// TIA Portal project "MiniProject_AziziFarid" (V16)

(* hardware
DEVICE "S71500/ET200MP station_1"  S7-1500 station
   slot 0: "Rail_0"  Rack  6ES7 590-1***0-0AA0
   slot 1: "AF_PLC_1 Distribution"  CPU 1512C-1 PN  6ES7 512-1CK00-0AB0  V2.6
      slot 3: "CPU display_1"  6ES7591-1AA00-0AA0
      slot 32768: "PROFINET interface_1"  X1
DEVICE "S71500/ET200MP station_2"  S7-1500 station
   slot 0: "Rail_0"  Rack  6ES7 590-1***0-0AA0
   slot 1: "AF_PLC_2 Joining"  CPU 1512C-1 PN  6ES7 512-1CK00-0AB0  V2.1
      slot 3: "CPU display_1"  6ES7591-1AA00-0AA0
      slot 32768: "PROFINET interface_1"  X1
DEVICE "S71500/ET200MP station_3"  S7-1500 station
   slot 0: "Rail_0"  Rack  6ES7 590-1***0-0AA0
   slot 1: "AF_PLC_3 Sorting"  CPU 1512C-1 PN  6ES7 512-1CK00-0AB0  V2.1
      slot 3: "CPU display_1"  6ES7591-1AA00-0AA0
      slot 32768: "PROFINET interface_1"  X1
DEVICE "GSD device_1"  GSD.Device.PN
   slot 0: "Rack"  Rack  V1.0
   slot 0: "CTEU-PN"  CTEU-PN  2201471
      slot 0: "CTEU-PN"  CTEU-PN
      slot 1: "PN-IO Interface"  PN-IO Interface
         slot 1: "Port 1"  Port 1
         slot 2: "Port 2"  Port 2
   slot 1: "Universal device 064DIO_1"  Universal device 064DIO
      slot 0: "Universal device 064DIO"  Universal device 064DIO
*)

// ===== PLC "AF_PLC_1 Distribution"  CPU 1512C-1 PN =====

VAR_GLOBAL   // PLC tag table "Default tag table"
   "SF1 START BTN" AT %I11.0 : Bool;
   "SF2 STOP BTN" AT %I11.1 : Bool;
   "SF4 KEY SWITCH" AT %I11.2 : Bool;
   "SF3 RESET BTN" AT %I11.3 : Bool;
   "G1BG1 SENSOR1" AT %I10.0 : Bool;
   "G1BG2 SENSOR2" AT %I10.1 : Bool;
   "G1BG3 SENSOR3" AT %I10.2 : Bool;
   "C2BG1 SLIDE RETRACT" AT %I10.4 : Bool;
   "C2BG2 SLIDE EXTEND" AT %I10.5 : Bool;
   "C2BG3 MAGAZINE EMPTY" AT %I10.6 : Bool;
   "PF1 START IND" AT %Q5.0 : Bool;
   "PF2 RESET IND" AT %Q5.1 : Bool;
   "PF3 IND Q1" AT %Q5.2 : Bool;
   "q4 XD4 STATION FREE" AT %Q5.4 : Bool;
   "q5 indLightGn" AT %Q5.5 : Bool;
   "q6 indLightYe" AT %Q5.6 : Bool;
   "q7 indLightRd" AT %Q5.7 : Bool;
   "G1BF1_A1 CONV FRWD" AT %Q4.0 : Bool;
   "G1BF1_A2 CONV BKWD" AT %Q4.1 : Bool;
   "G1MB1" AT %Q4.2 : Bool;
   "C2MB1" AT %Q4.4 : Bool;
   "System_Byte" AT %MB999 : Byte;
   "FirstScan" AT %M999.0 : Bool;
   "DiagStatusUpdate" AT %M999.1 : Bool;
   "AlwaysTRUE" AT %M999.2 : Bool;
   "AlwaysFALSE" AT %M999.3 : Bool;
   "Clock_Byte" AT %MB1000 : Byte;
   "Clock_10Hz" AT %M1000.0 : Bool;
   "Clock_5Hz" AT %M1000.1 : Bool;
   "Clock_2.5Hz" AT %M1000.2 : Bool;
   "Clock_2Hz" AT %M1000.3 : Bool;
   "Clock_1.25Hz" AT %M1000.4 : Bool;
   "Clock_1Hz" AT %M1000.5 : Bool;
   "Clock_0.625Hz" AT %M1000.6 : Bool;
   "Clock_0.5Hz" AT %M1000.7 : Bool;
   "xResetModules" AT %M200.0 : Bool;
   "xResetReadyModule1" AT %M200.1 : Bool;
   "xResetReadyModule2" AT %M200.2 : Bool;
   "xResetReadyModule3" AT %M200.3 : Bool;
   "xEnAutoMM" AT %M300.0 : Bool;
   "xDeactivateModules" AT %M200.6 : Bool;
   "xProcessBusyMM" AT %M200.7 : Bool;
   "xResetReadyMM" AT %M201.0 : Bool;
   "xNextStationFreeMM" AT %M201.1 : Bool;
   "xReadyModSM" AT %M201.2 : Bool;
   "xStartModuleSM" AT %M201.3 : Bool;
   "xMagEmptySM" AT %M201.4 : Bool;
   "xInitModules" AT %M201.5 : Bool;
   "PF4" AT %Q5.3 : Bool;
   "i7 XD7" AT %I11.7 : Bool;
   "i5 SF5" AT %I11.5 : Bool;
   "xResetReadyRFID_1" AT %M201.6 : Bool;
   "xMActivateModule1" AT %M201.7 : Bool;
   "xMEnAuto" AT %M400.7 : Bool;
   "xMStartProcess" AT %M300.2 : Bool;
   "xMProcessBusy" AT %M300.1 : Bool;
   "xMTP" AT %M203.0 : Bool;
   "xMTFR" AT %M203.1 : Bool;
   "xMG1BF1_A1" AT %M203.2 : Bool;
   "xM_MES_EnAuto" AT %M300.3 : Bool;
   "MWtest" AT %MW550 : Word;
   "bErrCodeMod1" AT %MB450 : Byte;
   "bErrCodeMod2" AT %MB451 : Byte;
   "bErrCodeMod3" AT %MB452 : Byte;
   "bErrCodeSeq" AT %MB453 : Byte;
   "bErrCodeOpMode" AT %MB454 : Byte;
   "Tag_1" AT %C2 : Counter;
   "i6 Jumper" AT %I11.6 : Bool;
   "Output" AT %M0.1 : Bool;
   "i4" AT %I11.4 : Bool;
   "Tag_2" AT %M0.0 : Bool;
   "Tag_3" AT %Q4.3 : Bool;
END_VAR

DATA_BLOCK "Dist_Block_DB"   // DB1
{ S7_Optimized_Access := 'TRUE' }
VERSION : 0.1
// stored: InstanceOfName Dist_Block
"Dist_Block"
BEGIN
END_DATA_BLOCK

// folder: System blocks/Program resources

DATA_BLOCK "IEC_Counter_0_DB"   // DB2
{ S7_Optimized_Access := 'TRUE' }
AUTHOR : Simatic
FAMILY : IEC
NAME : CNTR
VERSION : 1.0
// stored: InstanceOfName IEC_COUNTER
"IEC_COUNTER"
BEGIN
END_DATA_BLOCK

// folder: (top level)

FUNCTION_BLOCK "Dist_Block"   // FB2, GRAPH_PLUS
{ S7_Optimized_Access := 'TRUE' }
VERSION : 0.1
   VAR_INPUT
      OFF_SQ : Bool := false;   // Turn sequence off
      INIT_SQ : Bool := false;   // Set sequence to initial state
      ACK_EF : Bool := false;   // Acknowledge all errors and faults
      S_PREV : Bool := false;   // Output previous step in parameter S_NO
      S_NEXT : Bool := false;   // Indicate next step in parameter S_NO
      SW_AUTO : Bool := false;   // Automatic mode
      SW_TAP : Bool := false;   // Semiautomatic/switch with transition
      SW_TOP : Bool := false;   // Semiautomatic/ignore transition
      SW_MAN : Bool := false;   // Manual mode
      S_SEL : Int := 0;   // Select step to be output to S_NO
      S_ON : Bool := false;   // Activate step indicated in S_NO
      S_OFF : Bool := false;   // Deactivate step indicated S_NO
      T_PUSH : Bool := false;   // Enable transition to switch in semi automatic mode
   END_VAR
   VAR_OUTPUT
      S_NO : Int := 0;   // Step number
      S_MORE : Bool := false;   // More steps are available and can be shown in S_NO
      S_ACTIVE : Bool := false;   // Step indicated in S_NO is active
      ERR_FLT : Bool := false;   // Interlock or supervision group error
      AUTO_ON : Bool := false;   // Automatic mode is active
      TAP_ON : Bool := false;   // Semiautomatic mode/step with transition enabled
      TOP_ON : Bool := false;   // Semiautomatic mode/ignore transition enabled
      MAN_ON : Bool := false;   // Manual mode is active
   END_VAR
   VAR
      HMI_INFO : Array[0..8] of UInt;
      IF_PAR : G7_IfParPlus_V6;
      RT_DATA : G7_RTDataPlus_V6;   // Internal data area
      Trans1 : G7_TransitionPlus_V6;   // Transition structure
      Trans2 : G7_TransitionPlus_V6;   // Transition structure
      Trans3 : G7_TransitionPlus_V6;   // Transition structure
      Trans4 : G7_TransitionPlus_V6;   // Transition structure
      Trans5 : G7_TransitionPlus_V6;   // Transition structure
      Trans8 : G7_TransitionPlus_V6;   // Transition structure
      Trans9 : G7_TransitionPlus_V6;   // Transition structure
      Trans12 : G7_TransitionPlus_V6;   // Transition structure
      Trans13 : G7_TransitionPlus_V6;   // Transition structure
      Trans14 : G7_TransitionPlus_V6;   // Transition structure
      Step1 : G7_StepPlus_V6;   // Step structure
      Step2 : G7_StepPlus_V6;   // Step structure
      Step3 : G7_StepPlus_V6;   // Step structure
      Step4 : G7_StepPlus_V6;   // Step structure
      Step5 : G7_StepPlus_V6;   // Step structure
      Step8 : G7_StepPlus_V6;   // Step structure
      Step10 : G7_StepPlus_V6;   // Step structure
      Step11 : G7_StepPlus_V6;   // Step structure
      SINI : Array[0..1] of USInt;
      LSTT : Array[0..9] of USInt;
      ATAJ : Array[0..9] of USInt;
      ATAB : Array[0..9] of USInt;
      PSTT : Array[0..9] of USInt;
      NSTT : Array[0..9] of USInt;
      ASSJ : Array[0..7] of USInt;
      ASSB : Array[0..7] of USInt;
      PTTS : Array[0..7] of USInt;
      NTTS : Array[0..7] of USInt;
      SW_SQTS : Array[0..7] of USInt;
      SWITCH : Array[0..3] of USInt;
      TVX : Array[0..5] of USInt;
      TTX : Array[0..5] of USInt;
      TSX : Array[0..1] of USInt;
      S00X : Array[0..1] of USInt;
      SOFFX : Array[0..1] of USInt;
      SONX : Array[0..1] of USInt;
      SAX : Array[0..1] of USInt;
      SERRX : Array[0..8] of USInt;
      SMX : Array[0..8] of USInt;
      S0X : Array[0..8] of USInt;
      S1X : Array[0..8] of USInt;
      IL_ALARM_INST : Diag_Alarm;
      SUP_ALARM_INST : Diag_Alarm;
      STEP_TIME_ALARM_INST : Diag_Alarm;
      IEC_TIMER_INST : IEC_TIMER;
      TRANSACTION_FLAG : Bool := false;
   END_VAR
   // SINI[0] := 2;
   // LSTT[0] := 255;
   // LSTT[1] := 255;
   // LSTT[2] := 255;
   // ATAJ[1] := 1;
   // ATAJ[2] := 2;
   // ATAJ[3] := 3;
   // ATAB[1] := 1;
   // ATAB[2] := 2;
   // ATAB[3] := 7;
   // PSTT[1] := 1;
   // PSTT[2] := 2;
   // PSTT[3] := 3;
   // NSTT[0] := 1;
   // NSTT[1] := 2;
   // NSTT[2] := 3;
   // ASSJ[1] := 1;
   // ASSJ[2] := 2;
   // ASSJ[3] := 3;
   // ASSB[1] := 1;
   // ASSB[2] := 2;
   // ASSB[3] := 3;
   // PTTS[0] := 9;
   // PTTS[2] := 1;
   // PTTS[3] := 2;
   // NTTS[1] := 1;
   // NTTS[2] := 2;
   // NTTS[3] := 3;
   // TVX[0] := 16#1;
   // TTX[0] := 16#1;
   // TSX[0] := 16#1;
   // S00X[0] := 16#1;
   // SOFFX[0] := 16#1;
   // SONX[0] := 16#1;
   // SAX[0] := 16#1;
   // SERRX[0] := 16#1;
   // SMX[0] := 16#1;
   // S0X[0] := 16#1;
   // S1X[0] := 16#1;
   // ATAB[0] := 5;
   // LSTT[5] := 255;
   // ATAJ[4] := 4;
   // ATAJ[5] := 5;
   // ATAB[7] := 3;
   // NSTT[5] := 5;
   // ASSJ[4] := 4;
   // ASSB[4] := 4;
   // PTTS[4] := 3;
   // NTTS[4] := 4;
   // SW_SQTS[1] := 1;
   // SW_SQTS[2] := 1;
   // SW_SQTS[3] := 1;
   // SW_SQTS[4] := 2;
   // LSTT[3] := 255;
   // ATAJ[6] := 6;
   // ATAB[4] := 4;
   // PSTT[4] := 4;
   // NSTT[3] := 4;
   // ASSJ[5] := 5;
   // ASSB[5] := 5;
   // PTTS[5] := 5;
   // NTTS[6] := 8;
   // SW_SQTS[6] := 4;
   // LSTT[7] := 255;
   // ATAJ[7] := 7;
   // ATAB[6] := 6;
   // PSTT[7] := 3;
   // NSTT[7] := 6;
   // ASSJ[6] := 6;
   // ASSB[6] := 6;
   // PTTS[6] := 7;
   // NTTS[5] := 6;
   // LSTT[9] := 255;
   // ATAJ[8] := 8;
   // ATAJ[9] := 9;
   // ATAB[8] := 8;
   // ATAB[9] := 9;
   // PSTT[8] := 6;
   // PSTT[9] := 7;
   // ASSJ[7] := 7;
   // ASSB[7] := 7;
   // PTTS[7] := 255;
   // NTTS[7] := 9;
   // PSTT[6] := 5;
   // SW_SQTS[5] := 3;
BEGIN
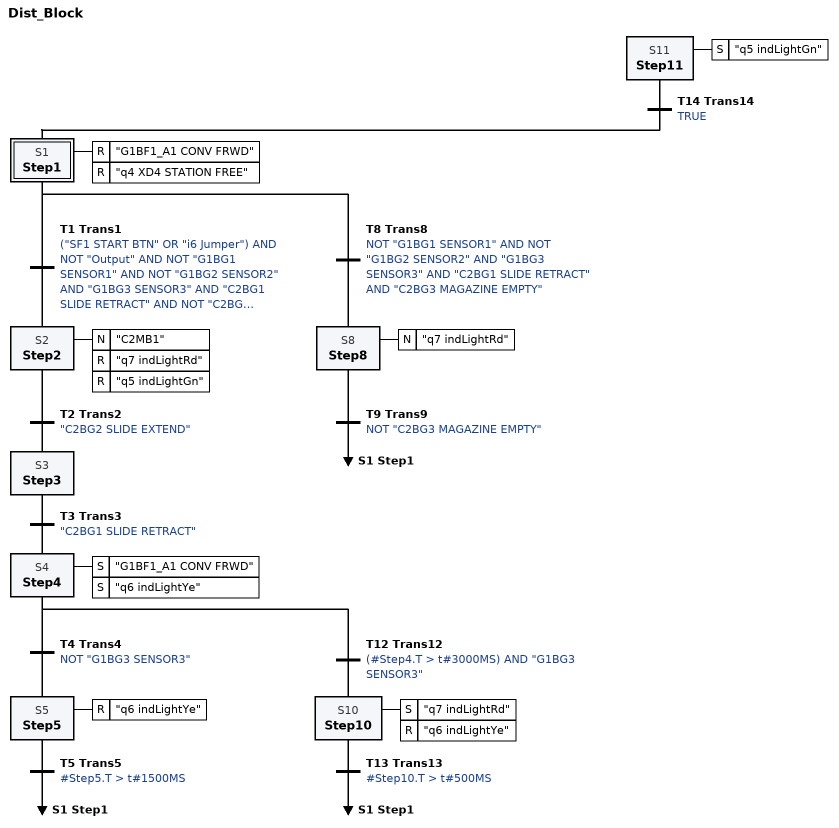
   // sequencer 1
   INITIAL_STEP Step1:   // S1, max time T#10S, warning time T#7S
              R    "G1BF1_A1 CONV FRWD"
              R    "q4 XD4 STATION FREE"
   END_STEP
   TRANSITION Trans1 FROM Step1 TO Step2   // T1
      := ("SF1 START BTN" OR "i6 Jumper") AND NOT "Output" AND NOT "G1BG1 SENSOR1" AND NOT "G1BG2 SENSOR2" AND "G1BG3 SENSOR3" AND "C2BG1 SLIDE RETRACT" AND NOT "C2BG3 MAGAZINE EMPTY";
   END_TRANSITION
   TRANSITION Trans8 FROM Step1 TO Step8   // T8
      := NOT "G1BG1 SENSOR1" AND NOT "G1BG2 SENSOR2" AND "G1BG3 SENSOR3" AND "C2BG1 SLIDE RETRACT" AND "C2BG3 MAGAZINE EMPTY";
   END_TRANSITION
   STEP Step2:   // S2, max time T#10S, warning time T#7S
              N    "C2MB1"
              R    "q7 indLightRd"
              R    "q5 indLightGn"
   END_STEP
   TRANSITION Trans2 FROM Step2 TO Step3   // T2
      := "C2BG2 SLIDE EXTEND";
   END_TRANSITION
   STEP Step3:   // S3, max time T#10S, warning time T#7S
   END_STEP
   TRANSITION Trans3 FROM Step3 TO Step4   // T3
      := "C2BG1 SLIDE RETRACT";
   END_TRANSITION
   STEP Step4:   // S4, max time T#10S, warning time T#7S
              S    "G1BF1_A1 CONV FRWD"
              S    "q6 indLightYe"
   END_STEP
   TRANSITION Trans4 FROM Step4 TO Step5   // T4
      := NOT "G1BG3 SENSOR3";
   END_TRANSITION
   TRANSITION Trans12 FROM Step4 TO Step10   // T12
      := (#Step4.T > t#3000MS) AND "G1BG3 SENSOR3";
   END_TRANSITION
   STEP Step8:   // S8, max time T#10S, warning time T#7S
              N    "q7 indLightRd"
   END_STEP
   TRANSITION Trans9 FROM Step8 TO Step1   // T9, jump
      := NOT "C2BG3 MAGAZINE EMPTY";
   END_TRANSITION
   STEP Step5:   // S5, max time T#10S, warning time T#7S
              R    "q6 indLightYe"
   END_STEP
   TRANSITION Trans5 FROM Step5 TO Step1   // T5, jump
      := #Step5.T > t#1500MS;
   END_TRANSITION
   STEP Step10:   // S10, max time T#10S, warning time T#7S
              S    "q7 indLightRd"
              R    "q6 indLightYe"
   END_STEP
   TRANSITION Trans13 FROM Step10 TO Step1   // T13, jump
      := #Step10.T > t#500MS;
   END_TRANSITION
   STEP Step11:   // S11, max time T#10S, warning time T#7S
              S    "q5 indLightGn"
   END_STEP
   TRANSITION Trans14 FROM Step11 TO Step1   // T14
      := TRUE;
   END_TRANSITION
END_FUNCTION_BLOCK

ORGANIZATION_BLOCK "Dist_Main"   // OB1, LAD, ProgramCycle
TITLE = "Main Program Sweep (Cycle)"
{ S7_Optimized_Access := 'TRUE' }
VERSION : 0.1
   VAR_INPUT
      Initial_Call : Bool;   // Initial call of this OB
      Remanence : Bool;   // =True, if remanent data are available
   END_VAR
BEGIN

REGION Network 1
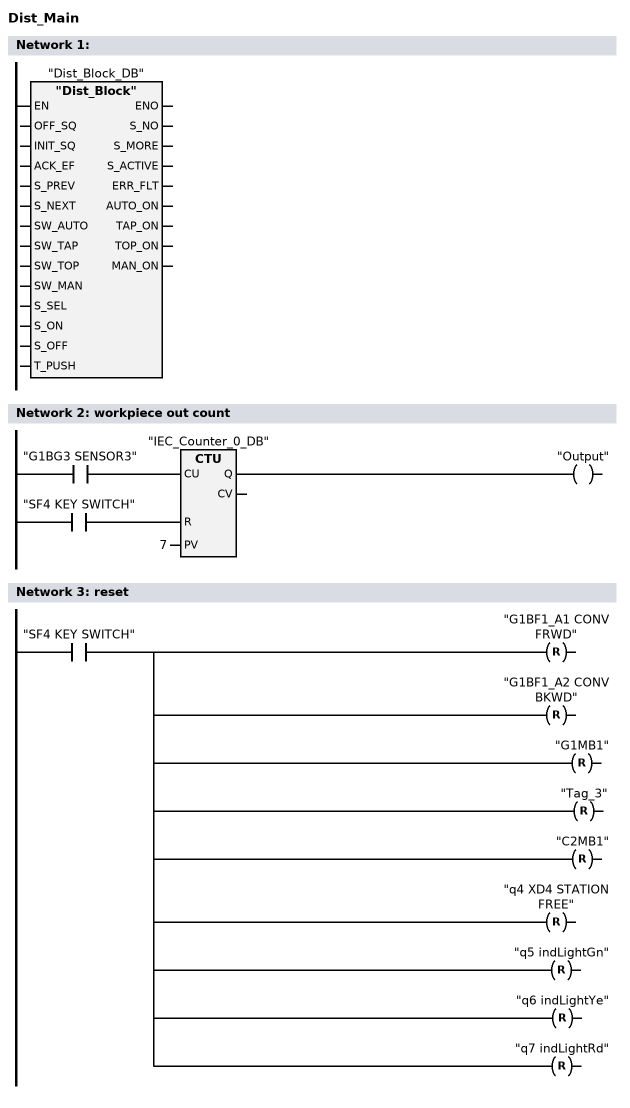
   RUNG wire#powerrail
      "Dist_Block_DB"(OFF_SQ :=, INIT_SQ :=, ACK_EF :=, S_PREV :=, S_NEXT :=, SW_AUTO :=, SW_TAP :=, SW_TOP :=, SW_MAN :=, S_SEL :=, S_ON :=, S_OFF :=, T_PUSH :=, S_NO =>, S_MORE =>, S_ACTIVE =>, ERR_FLT =>, AUTO_ON =>, TAP_ON =>, TOP_ON =>, MAN_ON =>)
   END_RUNG
   // the same network as SCL:
   "Dist_Block_DB"();   // "Dist_Block"
END_REGION

REGION Network 2: workpiece out count
   "IEC_Counter_0_DB".CTU(CU := "G1BG3 SENSOR3", R := "SF4 KEY SWITCH", PV := 7);
   "Output" := "IEC_Counter_0_DB".Q;
END_REGION

REGION Network 3: reset
   RUNG wire#powerrail
      Contact( "SF4 KEY SWITCH" )
      wire#w1
      R_Coil( "G1BF1_A1 CONV FRWD" )
   END_RUNG
   RUNG wire#w1
      R_Coil( "G1BF1_A2 CONV BKWD" )
   END_RUNG
   RUNG wire#w1
      R_Coil( "G1MB1" )
   END_RUNG
   RUNG wire#w1
      R_Coil( "Tag_3" )
   END_RUNG
   RUNG wire#w1
      R_Coil( "C2MB1" )
   END_RUNG
   RUNG wire#w1
      R_Coil( "q4 XD4 STATION FREE" )
   END_RUNG
   RUNG wire#w1
      R_Coil( "q5 indLightGn" )
   END_RUNG
   RUNG wire#w1
      R_Coil( "q6 indLightYe" )
   END_RUNG
   RUNG wire#w1
      R_Coil( "q7 indLightRd" )
   END_RUNG
   // the same network as SCL:
   IF "SF4 KEY SWITCH" THEN
       "G1BF1_A1 CONV FRWD" := FALSE;
       "G1BF1_A2 CONV BKWD" := FALSE;
       "G1MB1" := FALSE;
       "Tag_3" := FALSE;
       "C2MB1" := FALSE;
       "q4 XD4 STATION FREE" := FALSE;
       "q5 indLightGn" := FALSE;
       "q6 indLightYe" := FALSE;
       "q7 indLightRd" := FALSE;
   END_IF;
END_REGION
END_ORGANIZATION_BLOCK

// ===== PLC "AF_PLC_2 Joining"  CPU 1512C-1 PN =====

VAR_GLOBAL   // PLC tag table "Default tag table"
   "G1BG1 (diffuse 1 - depan)" AT %I10.0 : Bool;
   "G1BG2 (diffuse 2 - tengah)" AT %I10.1 : Bool;
   "G1MB1 (sep)" AT %Q4.2 : Bool;
   "G1MB2 (stopper)" AT %Q4.3 : Bool;
   "G1KF1-1 conv fwd" AT %Q4.0 : Bool;
   "G2BG3" AT %I10.6 : Bool;
   "G1KF1-2 conv bwd" AT %Q4.1 : Bool;
   "G1BG3 (through beam - hujung)" AT %I10.2 : Bool;
   "G1BG4 (distance)" AT %I10.3 : Bool;
   "G2KF1-1 conv fwd" AT %Q4.4 : Bool;
   "G2KF1-2 conv bwd" AT %Q4.5 : Bool;
   "G2BG1 (diffuse - capping)" AT %I10.4 : Bool;
   "SF1 (start btn)" AT %I11.0 : Bool;
   "SF2 (stop btn)" AT %I11.1 : Bool;
   "G3BG1 (sensor_arm_masuk)" AT %I126.0 : Bool;
   "G3BG2 (sensor_arm_keluar)" AT %I126.1 : Bool;
   "G3BG3 (sensor_arm_naik)" AT %I126.2 : Bool;
   "G3BP1 (sensor_sedut)" AT %I126.3 : Bool;
   "G3MB1 P1 (arm_keluar)" AT %Q128.1 : Bool;
   "G3MB2 P0 (arm_masuk)" AT %Q128.0 : Bool;
   "G3MB3 (arm_turunH_naikL)" AT %Q128.2 : Bool;
   "G3MB4 (sedut)" AT %Q128.3 : Bool;
   "SF3" AT %I11.2 : Bool;
   "SF4" AT %I11.3 : Bool;
   "i5" AT %I11.5 : Bool;
   "i6" AT %I11.6 : Bool;
   "i7" AT %I11.7 : Bool;
   "PF1" AT %I12.0 : Bool;
   "PF2" AT %I12.1 : Bool;
   "XPROCESSBUSY" AT %M0.0 : Bool;
   "i4 Jumper" AT %I11.4 : Bool;
   "output1" AT %M0.1 : Bool;
   "output2" AT %M0.2 : Bool;
   "q4" AT %Q5.4 : Bool;
   "q5" AT %Q5.5 : Bool;
   "q6" AT %Q5.6 : Bool;
   "q7" AT %Q5.7 : Bool;
END_VAR

DATA_BLOCK "Joining_Block_DB"   // DB1
{ S7_Optimized_Access := 'TRUE' }
VERSION : 0.1
// stored: InstanceOfName Joining_Block
"Joining_Block"
BEGIN
END_DATA_BLOCK

// folder: System blocks/Program resources

DATA_BLOCK "IEC_Counter_0_DB"   // DB2
{ S7_Optimized_Access := 'TRUE' }
AUTHOR : Simatic
FAMILY : IEC
NAME : CNTR
VERSION : 1.0
// stored: InstanceOfName IEC_COUNTER
"IEC_COUNTER"
BEGIN
END_DATA_BLOCK

DATA_BLOCK "IEC_Counter_0_DB_1"   // DB3
{ S7_Optimized_Access := 'TRUE' }
AUTHOR : Simatic
FAMILY : IEC
NAME : CNTR
VERSION : 1.0
// stored: InstanceOfName IEC_COUNTER
"IEC_COUNTER"
BEGIN
END_DATA_BLOCK

// folder: (top level)

FUNCTION_BLOCK "Joining_Block"   // FB1, GRAPH_PLUS
{ S7_Optimized_Access := 'TRUE' }
VERSION : 0.1
   VAR_INPUT
      OFF_SQ : Bool := false;   // Turn sequence off
      INIT_SQ : Bool := false;   // Set sequence to initial state
      ACK_EF : Bool := false;   // Acknowledge all errors and faults
      S_PREV : Bool := false;   // Output previous step in parameter S_NO
      S_NEXT : Bool := false;   // Indicate next step in parameter S_NO
      SW_AUTO : Bool := false;   // Automatic mode
      SW_TAP : Bool := false;   // Semiautomatic/switch with transition
      SW_TOP : Bool := false;   // Semiautomatic/ignore transition
      SW_MAN : Bool := false;   // Manual mode
      S_SEL : Int := 0;   // Select step to be output to S_NO
      S_ON : Bool := false;   // Activate step indicated in S_NO
      S_OFF : Bool := false;   // Deactivate step indicated S_NO
      T_PUSH : Bool := false;   // Enable transition to switch in semi automatic mode
   END_VAR
   VAR_OUTPUT
      S_NO : Int := 0;   // Step number
      S_MORE : Bool := false;   // More steps are available and can be shown in S_NO
      S_ACTIVE : Bool := false;   // Step indicated in S_NO is active
      ERR_FLT : Bool := false;   // Interlock or supervision group error
      AUTO_ON : Bool := false;   // Automatic mode is active
      TAP_ON : Bool := false;   // Semiautomatic mode/step with transition enabled
      TOP_ON : Bool := false;   // Semiautomatic mode/ignore transition enabled
      MAN_ON : Bool := false;   // Manual mode is active
   END_VAR
   VAR
      HMI_INFO : Array[0..8] of UInt;
      IF_PAR : G7_IfParPlus_V6;
      RT_DATA : G7_RTDataPlus_V6;   // Internal data area
      Trans1 : G7_TransitionPlus_V6;   // Transition structure
      Trans2 : G7_TransitionPlus_V6;   // Transition structure
      Trans3 : G7_TransitionPlus_V6;   // Transition structure
      Trans4 : G7_TransitionPlus_V6;   // Transition structure
      Trans5 : G7_TransitionPlus_V6;   // Transition structure
      Trans6 : G7_TransitionPlus_V6;   // Transition structure
      Trans7 : G7_TransitionPlus_V6;   // Transition structure
      Trans8 : G7_TransitionPlus_V6;   // Transition structure
      Trans9 : G7_TransitionPlus_V6;   // Transition structure
      Trans10 : G7_TransitionPlus_V6;   // Transition structure
      Trans11 : G7_TransitionPlus_V6;   // Transition structure
      Trans12 : G7_TransitionPlus_V6;   // Transition structure
      Trans13 : G7_TransitionPlus_V6;   // Transition structure
      Trans14 : G7_TransitionPlus_V6;   // Transition structure
      Trans15 : G7_TransitionPlus_V6;   // Transition structure
      Trans16 : G7_TransitionPlus_V6;   // Transition structure
      Trans17 : G7_TransitionPlus_V6;   // Transition structure
      Trans18 : G7_TransitionPlus_V6;   // Transition structure
      Trans19 : G7_TransitionPlus_V6;   // Transition structure
      Trans25 : G7_TransitionPlus_V6;   // Transition structure
      Trans26 : G7_TransitionPlus_V6;   // Transition structure
      Step1 : G7_StepPlus_V6;   // Step structure
      Step2 : G7_StepPlus_V6;   // Step structure
      Step3 : G7_StepPlus_V6;   // Step structure
      Step4 : G7_StepPlus_V6;   // Step structure
      Step5 : G7_StepPlus_V6;   // Step structure
      Step6 : G7_StepPlus_V6;   // Step structure
      Step8 : G7_StepPlus_V6;   // Step structure
      Step9 : G7_StepPlus_V6;   // Step structure
      Step10 : G7_StepPlus_V6;   // Step structure
      Step11 : G7_StepPlus_V6;   // Step structure
      Step12 : G7_StepPlus_V6;   // Step structure
      Step13 : G7_StepPlus_V6;   // Step structure
      Step14 : G7_StepPlus_V6;   // Step structure
      Step15 : G7_StepPlus_V6;   // Step structure
      Step16 : G7_StepPlus_V6;   // Step structure
      Step17 : G7_StepPlus_V6;   // Step structure
      Step18 : G7_StepPlus_V6;   // Step structure
      Step23 : G7_StepPlus_V6;   // Step structure
      Step24 : G7_StepPlus_V6;   // Step structure
      SINI : Array[0..1] of USInt;
      LSTT : Array[0..20] of USInt;
      ATAJ : Array[0..20] of USInt;
      ATAB : Array[0..20] of USInt;
      PSTT : Array[0..20] of USInt;
      NSTT : Array[0..20] of USInt;
      ASSJ : Array[0..18] of USInt;
      ASSB : Array[0..18] of USInt;
      PTTS : Array[0..18] of USInt;
      NTTS : Array[0..18] of USInt;
      SW_SQTS : Array[0..18] of USInt;
      SWITCH : Array[0..3] of USInt;
      TVX : Array[0..5] of USInt;
      TTX : Array[0..5] of USInt;
      TSX : Array[0..1] of USInt;
      S00X : Array[0..1] of USInt;
      SOFFX : Array[0..1] of USInt;
      SONX : Array[0..1] of USInt;
      SAX : Array[0..1] of USInt;
      SERRX : Array[0..19] of USInt;
      SMX : Array[0..19] of USInt;
      S0X : Array[0..19] of USInt;
      S1X : Array[0..19] of USInt;
      IL_ALARM_INST : Diag_Alarm;
      SUP_ALARM_INST : Diag_Alarm;
      STEP_TIME_ALARM_INST : Diag_Alarm;
      IEC_TIMER_INST : IEC_TIMER;
      TRANSACTION_FLAG : Bool := false;
   END_VAR
   // SINI[0] := 2;
   // LSTT[0] := 255;
   // LSTT[1] := 255;
   // LSTT[2] := 255;
   // LSTT[3] := 255;
   // LSTT[4] := 255;
   // LSTT[5] := 255;
   // LSTT[6] := 255;
   // LSTT[9] := 255;
   // ATAJ[1] := 1;
   // ATAJ[2] := 2;
   // ATAJ[3] := 3;
   // ATAJ[4] := 4;
   // ATAJ[5] := 5;
   // ATAJ[6] := 6;
   // ATAJ[7] := 7;
   // ATAJ[8] := 8;
   // ATAB[1] := 1;
   // ATAB[2] := 2;
   // ATAB[3] := 6;
   // ATAB[4] := 4;
   // ATAB[5] := 5;
   // ATAB[6] := 3;
   // ATAB[7] := 7;
   // ATAB[8] := 8;
   // PSTT[1] := 1;
   // PSTT[2] := 2;
   // PSTT[3] := 3;
   // PSTT[4] := 4;
   // PSTT[5] := 5;
   // PSTT[6] := 3;
   // PSTT[7] := 6;
   // PSTT[8] := 7;
   // NSTT[0] := 15;
   // NSTT[1] := 2;
   // NSTT[2] := 3;
   // NSTT[3] := 4;
   // NSTT[4] := 8;
   // NSTT[5] := 7;
   // NSTT[6] := 6;
   // NSTT[9] := 9;
   // ASSJ[1] := 1;
   // ASSJ[2] := 2;
   // ASSJ[3] := 3;
   // ASSJ[4] := 4;
   // ASSJ[5] := 5;
   // ASSJ[6] := 6;
   // ASSJ[7] := 7;
   // ASSB[1] := 1;
   // ASSB[2] := 2;
   // ASSB[3] := 3;
   // ASSB[4] := 4;
   // ASSB[5] := 5;
   // ASSB[6] := 6;
   // ASSB[7] := 7;
   // PTTS[0] := 255;
   // PTTS[2] := 1;
   // PTTS[3] := 2;
   // PTTS[4] := 3;
   // PTTS[5] := 14;
   // PTTS[6] := 6;
   // PTTS[7] := 5;
   // NTTS[1] := 1;
   // NTTS[2] := 2;
   // NTTS[3] := 3;
   // NTTS[4] := 4;
   // NTTS[5] := 5;
   // NTTS[6] := 7;
   // NTTS[7] := 8;
   // SW_SQTS[4] := 1;
   // SW_SQTS[5] := 2;
   // SW_SQTS[6] := 3;
   // SW_SQTS[7] := 2;
   // TVX[0] := 16#1;
   // TTX[0] := 16#1;
   // TSX[0] := 16#1;
   // S00X[0] := 16#1;
   // SOFFX[0] := 16#1;
   // SONX[0] := 16#1;
   // SAX[0] := 16#1;
   // SERRX[0] := 16#1;
   // SMX[0] := 16#1;
   // S0X[0] := 16#1;
   // S1X[0] := 16#1;
   // LSTT[10] := 255;
   // LSTT[11] := 255;
   // LSTT[12] := 255;
   // LSTT[13] := 255;
   // LSTT[14] := 255;
   // ATAJ[9] := 9;
   // ATAJ[10] := 10;
   // ATAJ[11] := 11;
   // ATAJ[12] := 12;
   // ATAJ[13] := 13;
   // ATAJ[14] := 14;
   // ATAB[9] := 9;
   // ATAB[10] := 17;
   // ATAB[11] := 11;
   // ATAB[12] := 12;
   // ATAB[13] := 13;
   // ATAB[14] := 14;
   // PSTT[9] := 8;
   // PSTT[10] := 9;
   // PSTT[11] := 10;
   // PSTT[12] := 11;
   // PSTT[13] := 12;
   // PSTT[14] := 13;
   // NSTT[10] := 10;
   // NSTT[11] := 11;
   // NSTT[12] := 12;
   // NSTT[13] := 13;
   // NSTT[14] := 5;
   // ASSJ[8] := 8;
   // ASSJ[9] := 9;
   // ASSJ[10] := 10;
   // ASSJ[11] := 11;
   // ASSJ[12] := 12;
   // ASSJ[13] := 13;
   // ASSB[8] := 8;
   // ASSB[9] := 9;
   // ASSB[10] := 10;
   // ASSB[11] := 11;
   // ASSB[12] := 12;
   // ASSB[13] := 13;
   // PTTS[8] := 4;
   // PTTS[9] := 9;
   // PTTS[10] := 10;
   // PTTS[11] := 11;
   // PTTS[12] := 12;
   // PTTS[13] := 13;
   // NTTS[8] := 9;
   // NTTS[9] := 10;
   // NTTS[10] := 11;
   // NTTS[11] := 12;
   // NTTS[12] := 13;
   // NTTS[13] := 14;
   // SW_SQTS[8] := 1;
   // SW_SQTS[9] := 1;
   // SW_SQTS[10] := 2;
   // SW_SQTS[11] := 2;
   // SW_SQTS[12] := 2;
   // SW_SQTS[13] := 2;
   // LSTT[7] := 255;
   // ATAJ[15] := 15;
   // ATAB[15] := 15;
   // PSTT[15] := 14;
   // NSTT[7] := 14;
   // ASSJ[14] := 14;
   // ASSB[14] := 14;
   // PTTS[14] := 7;
   // NTTS[14] := 15;
   // SW_SQTS[14] := 3;
   // LSTT[16] := 255;
   // ATAJ[16] := 16;
   // ATAB[16] := 16;
   // PSTT[16] := 15;
   // NSTT[16] := 1;
   // ASSJ[15] := 15;
   // ASSB[15] := 15;
   // PTTS[1] := 16;
   // NTTS[15] := 16;
   // LSTT[17] := 255;
   // LSTT[18] := 255;
   // ATAJ[17] := 17;
   // ATAJ[18] := 18;
   // ATAB[17] := 10;
   // ATAB[18] := 18;
   // PSTT[17] := 9;
   // PSTT[18] := 16;
   // NSTT[17] := 16;
   // NSTT[18] := 18;
   // ASSJ[16] := 16;
   // ASSB[16] := 16;
   // PTTS[16] := 17;
   // NTTS[16] := 18;
   // SW_SQTS[16] := 4;
   // LSTT[20] := 255;
   // ATAJ[19] := 19;
   // ATAJ[20] := 20;
   // ATAB[19] := 19;
   // ATAB[20] := 20;
   // PSTT[19] := 17;
   // PSTT[20] := 18;
   // NSTT[20] := 17;
   // ASSJ[17] := 17;
   // ASSJ[18] := 18;
   // ASSB[17] := 17;
   // ASSB[18] := 18;
   // PTTS[17] := 20;
   // PTTS[18] := 18;
   // NTTS[17] := 19;
   // NTTS[18] := 20;
   // SW_SQTS[17] := 4;
   // SW_SQTS[18] := 4;
BEGIN
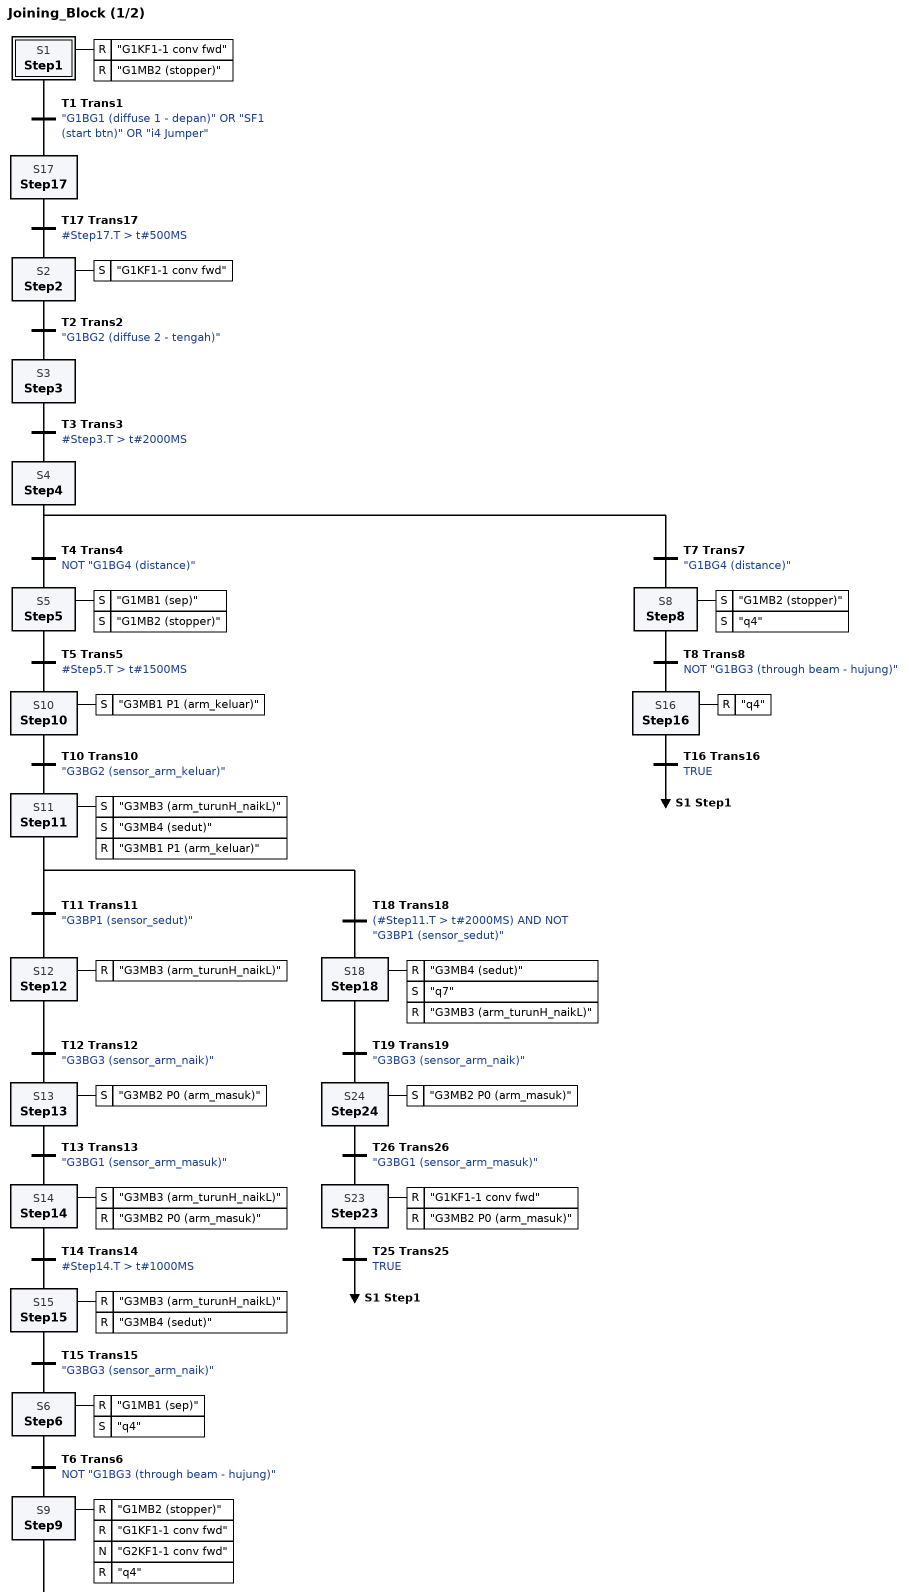
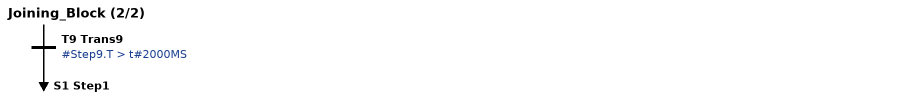
   // sequencer 1
   INITIAL_STEP Step1:   // S1, max time T#10S, warning time T#7S
              R    "G1KF1-1 conv fwd"
              R    "G1MB2 (stopper)"
   END_STEP
   TRANSITION Trans1 FROM Step1 TO Step17   // T1
      := "G1BG1 (diffuse 1 - depan)" OR "SF1 (start btn)" OR "i4 Jumper";
   END_TRANSITION
   STEP Step2:   // S2, max time T#10S, warning time T#7S
              S    "G1KF1-1 conv fwd"
   END_STEP
   TRANSITION Trans2 FROM Step2 TO Step3   // T2
      := "G1BG2 (diffuse 2 - tengah)";
   END_TRANSITION
   STEP Step3:   // S3, max time T#10S, warning time T#7S
   END_STEP
   TRANSITION Trans3 FROM Step3 TO Step4   // T3
      := #Step3.T > t#2000MS;
   END_TRANSITION
   STEP Step4:   // S4, max time T#10S, warning time T#7S
   END_STEP
   TRANSITION Trans4 FROM Step4 TO Step5   // T4
      := NOT "G1BG4 (distance)";
   END_TRANSITION
   TRANSITION Trans7 FROM Step4 TO Step8   // T7: Terbalik
      := "G1BG4 (distance)";
   END_TRANSITION
   STEP Step5:   // S5, max time T#10S, warning time T#7S
              S    "G1MB1 (sep)"
              S    "G1MB2 (stopper)"
   END_STEP
   TRANSITION Trans5 FROM Step5 TO Step10   // T5
      := #Step5.T > t#1500MS;
   END_TRANSITION
   STEP Step6:   // S6, max time T#10S, warning time T#7S
              R    "G1MB1 (sep)"
              S    "q4"
   END_STEP
   TRANSITION Trans6 FROM Step6 TO Step9   // T6
      := NOT "G1BG3 (through beam - hujung)";
   END_TRANSITION
   STEP Step8:   // S8, max time T#10S, warning time T#7S
              S    "G1MB2 (stopper)"
              S    "q4"
   END_STEP
   TRANSITION Trans8 FROM Step8 TO Step16   // T8
      := NOT "G1BG3 (through beam - hujung)";
   END_TRANSITION
   STEP Step9:   // S9, max time T#10S, warning time T#7S
              R    "G1MB2 (stopper)"
              R    "G1KF1-1 conv fwd"
              N    "G2KF1-1 conv fwd"
              R    "q4"
   END_STEP
   TRANSITION Trans9 FROM Step9 TO Step1   // T9, jump
      := #Step9.T > t#2000MS;
   END_TRANSITION
   STEP Step10:   // S10, max time T#10S, warning time T#7S
              S    "G3MB1 P1 (arm_keluar)"
   END_STEP
   TRANSITION Trans10 FROM Step10 TO Step11   // T10
      := "G3BG2 (sensor_arm_keluar)";
   END_TRANSITION
   STEP Step11:   // S11, max time T#10S, warning time T#7S
              S    "G3MB3 (arm_turunH_naikL)"
              S    "G3MB4 (sedut)"
              R    "G3MB1 P1 (arm_keluar)"
   END_STEP
   TRANSITION Trans11 FROM Step11 TO Step12   // T11
      := "G3BP1 (sensor_sedut)";
   END_TRANSITION
   TRANSITION Trans18 FROM Step11 TO Step18   // T18
      := (#Step11.T > t#2000MS) AND NOT "G3BP1 (sensor_sedut)";
   END_TRANSITION
   STEP Step12:   // S12, max time T#10S, warning time T#7S
              R    "G3MB3 (arm_turunH_naikL)"
   END_STEP
   TRANSITION Trans12 FROM Step12 TO Step13   // T12
      := "G3BG3 (sensor_arm_naik)";
   END_TRANSITION
   STEP Step13:   // S13, max time T#10S, warning time T#7S
      // undo Arm
              S    "G3MB2 P0 (arm_masuk)"
   END_STEP
   TRANSITION Trans13 FROM Step13 TO Step14   // T13
      := "G3BG1 (sensor_arm_masuk)";
   END_TRANSITION
   STEP Step14:   // S14, max time T#10S, warning time T#7S
      // turun Arm
              S    "G3MB3 (arm_turunH_naikL)"
              R    "G3MB2 P0 (arm_masuk)"
   END_STEP
   TRANSITION Trans14 FROM Step14 TO Step15   // T14
      := #Step14.T > t#1000MS;
   END_TRANSITION
   STEP Step15:   // S15, max time T#10S, warning time T#7S
      // pasang Cap
              R    "G3MB3 (arm_turunH_naikL)"
              R    "G3MB4 (sedut)"
   END_STEP
   TRANSITION Trans15 FROM Step15 TO Step6   // T15
      := "G3BG3 (sensor_arm_naik)";
   END_TRANSITION
   STEP Step16:   // S16, max time T#10S, warning time T#7S
              R    "q4"
   END_STEP
   TRANSITION Trans16 FROM Step16 TO Step1   // T16, jump
      := TRUE;
   END_TRANSITION
   STEP Step17:   // S17, max time T#10S, warning time T#7S
   END_STEP
   TRANSITION Trans17 FROM Step17 TO Step2   // T17
      := #Step17.T > t#500MS;
   END_TRANSITION
   STEP Step18:   // S18, max time T#10S, warning time T#7S
      // Lampu Merah
              R    "G3MB4 (sedut)"
              S    "q7"
              R    "G3MB3 (arm_turunH_naikL)"
   END_STEP
   TRANSITION Trans19 FROM Step18 TO Step24   // T19
      := "G3BG3 (sensor_arm_naik)";
   END_TRANSITION
   STEP Step24:   // S24, max time T#10S, warning time T#7S
              S    "G3MB2 P0 (arm_masuk)"
   END_STEP
   TRANSITION Trans26 FROM Step24 TO Step23   // T26
      := "G3BG1 (sensor_arm_masuk)";
   END_TRANSITION
   STEP Step23:   // S23, max time T#10S, warning time T#7S
              R    "G1KF1-1 conv fwd"
              R    "G3MB2 P0 (arm_masuk)"
   END_STEP
   TRANSITION Trans25 FROM Step23 TO Step1   // T25, jump
      := TRUE;
   END_TRANSITION
END_FUNCTION_BLOCK

ORGANIZATION_BLOCK "Joining_Main"   // OB1, LAD, ProgramCycle
TITLE = "Main Program Sweep (Cycle)"
{ S7_Optimized_Access := 'TRUE' }
VERSION : 0.1
   VAR_INPUT
      Initial_Call : Bool;   // Initial call of this OB
      Remanence : Bool;   // =True, if remanent data are available
   END_VAR
BEGIN

REGION Network 1
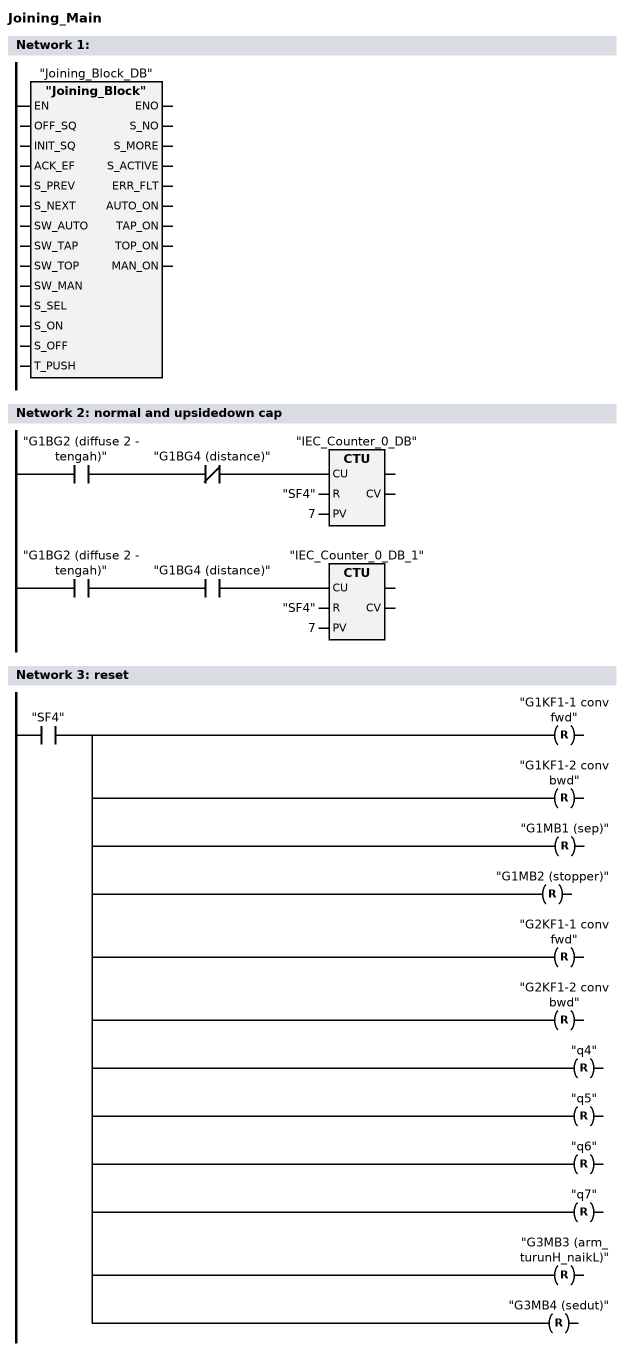
   RUNG wire#powerrail
      "Joining_Block_DB"(OFF_SQ :=, INIT_SQ :=, ACK_EF :=, S_PREV :=, S_NEXT :=, SW_AUTO :=, SW_TAP :=, SW_TOP :=, SW_MAN :=, S_SEL :=, S_ON :=, S_OFF :=, T_PUSH :=, S_NO =>, S_MORE =>, S_ACTIVE =>, ERR_FLT =>, AUTO_ON =>, TAP_ON =>, TOP_ON =>, MAN_ON =>)
   END_RUNG
   // the same network as SCL:
   "Joining_Block_DB"();   // "Joining_Block"
END_REGION

REGION Network 2: normal and upsidedown cap
   "IEC_Counter_0_DB".CTU(CU := "G1BG2 (diffuse 2 - tengah)" AND NOT "G1BG4 (distance)", R := "SF4", PV := 7);
   "IEC_Counter_0_DB_1".CTU(CU := "G1BG2 (diffuse 2 - tengah)" AND "G1BG4 (distance)", R := "SF4", PV := 7);
END_REGION

REGION Network 3: reset
   RUNG wire#powerrail
      Contact( "SF4" )
      wire#w1
      R_Coil( "G1KF1-1 conv fwd" )
   END_RUNG
   RUNG wire#w1
      R_Coil( "G1KF1-2 conv bwd" )
   END_RUNG
   RUNG wire#w1
      R_Coil( "G1MB1 (sep)" )
   END_RUNG
   RUNG wire#w1
      R_Coil( "G1MB2 (stopper)" )
   END_RUNG
   RUNG wire#w1
      R_Coil( "G2KF1-1 conv fwd" )
   END_RUNG
   RUNG wire#w1
      R_Coil( "G2KF1-2 conv bwd" )
   END_RUNG
   RUNG wire#w1
      R_Coil( "q4" )
   END_RUNG
   RUNG wire#w1
      R_Coil( "q5" )
   END_RUNG
   RUNG wire#w1
      R_Coil( "q6" )
   END_RUNG
   RUNG wire#w1
      R_Coil( "q7" )
   END_RUNG
   RUNG wire#w1
      R_Coil( "G3MB3 (arm_turunH_naikL)" )
   END_RUNG
   RUNG wire#w1
      R_Coil( "G3MB4 (sedut)" )
   END_RUNG
   // the same network as SCL:
   IF "SF4" THEN
       "G1KF1-1 conv fwd" := FALSE;
       "G1KF1-2 conv bwd" := FALSE;
       "G1MB1 (sep)" := FALSE;
       "G1MB2 (stopper)" := FALSE;
       "G2KF1-1 conv fwd" := FALSE;
       "G2KF1-2 conv bwd" := FALSE;
       "q4" := FALSE;
       "q5" := FALSE;
       "q6" := FALSE;
       "q7" := FALSE;
       "G3MB3 (arm_turunH_naikL)" := FALSE;
       "G3MB4 (sedut)" := FALSE;
   END_IF;
END_REGION
END_ORGANIZATION_BLOCK

// ===== PLC "AF_PLC_3 Sorting"  CPU 1512C-1 PN =====

VAR_GLOBAL   // PLC tag table "Default tag table"
   "SF1_START_BT" AT %I11.0 : Bool;
   "SF2_STOP_BT" AT %I11.1 : Bool;
   "SF4_KS MAN_AUTO" AT %I11.2 : Bool;
   "PF1_START INDI_LIGHT" AT %Q5.0 : Bool;
   "PF2_RESET INDI_LIGHT" AT %Q5.1 : Bool;
   "PF3(Q1)_INDI_LIGHT Q1" AT %Q5.2 : Bool;
   "PF4_INDI_LIGHT Q2" AT %Q5.3 : Bool;
   "B1BG1_FORK LIGHT BAR" AT %I10.4 : Bool;
   "B1BG2_RETRO LIGHT SENSOR" AT %I10.5 : Bool;
   "B1BG3_INDUC PROXI SENSOR" AT %I10.6 : Bool;
   "G1BG1_WP START" AT %I10.0 : Bool;
   "G1BG2_SEPARATOR 1 EXTRACT" AT %I10.1 : Bool;
   "G1BG4_SEPARATOR 2 EXTRACT" AT %I10.3 : Bool;
   "G1KF1_CONVEY MOTOR FOWD" AT %Q4.0 : Bool;
   "G1MB1_EXTEND SEPARATOR 1" AT %Q4.1 : Bool;
   "G1MB2_EXTEND SEPARATOR 2" AT %Q4.2 : Bool;
   "G1BG3_SENSOR SLIDE" AT %I10.2 : Bool;
   "G1MB3_RETRACT GATE" AT %Q4.3 : Bool;
   "q4 XD4_STATION FREE" AT %Q5.4 : Bool;
   "q5" AT %Q5.5 : Bool;
   "q6" AT %Q5.6 : Bool;
   "q7" AT %Q5.7 : Bool;
   "i4 Jumper" AT %I11.4 : Bool;
   "i5" AT %I11.5 : Bool;
   "i6 STATION_BUSY" AT %I11.6 : Bool;
   "i7" AT %I11.7 : Bool;
END_VAR

DATA_BLOCK "Sorting_Block_DB"   // DB1
{ S7_Optimized_Access := 'TRUE' }
VERSION : 0.1
// stored: InstanceOfName Sorting_Block
"Sorting_Block"
BEGIN
END_DATA_BLOCK

// folder: System blocks/Program resources

DATA_BLOCK "IEC_Counter_0_DB"   // DB2
{ S7_Optimized_Access := 'TRUE' }
AUTHOR : Simatic
FAMILY : IEC
NAME : CNTR
VERSION : 1.0
// stored: InstanceOfName IEC_COUNTER
"IEC_COUNTER"
BEGIN
END_DATA_BLOCK

DATA_BLOCK "IEC_Counter_0_DB_1"   // DB3
{ S7_Optimized_Access := 'TRUE' }
AUTHOR : Simatic
FAMILY : IEC
NAME : CNTR
VERSION : 1.0
// stored: InstanceOfName IEC_COUNTER
"IEC_COUNTER"
BEGIN
END_DATA_BLOCK

DATA_BLOCK "IEC_Counter_0_DB_2"   // DB4
{ S7_Optimized_Access := 'TRUE' }
AUTHOR : Simatic
FAMILY : IEC
NAME : CNTR
VERSION : 1.0
// stored: InstanceOfName IEC_COUNTER
"IEC_COUNTER"
BEGIN
END_DATA_BLOCK

// folder: (top level)

FUNCTION_BLOCK "Sorting_Block"   // FB3, GRAPH_PLUS
{ S7_Optimized_Access := 'TRUE' }
VERSION : 0.1
   VAR_INPUT
      OFF_SQ : Bool := false;   // Turn sequence off
      INIT_SQ : Bool := false;   // Set sequence to initial state
      ACK_EF : Bool := false;   // Acknowledge all errors and faults
      S_PREV : Bool := false;   // Output previous step in parameter S_NO
      S_NEXT : Bool := false;   // Indicate next step in parameter S_NO
      SW_AUTO : Bool := false;   // Automatic mode
      SW_TAP : Bool := false;   // Semiautomatic/switch with transition
      SW_TOP : Bool := false;   // Semiautomatic/ignore transition
      SW_MAN : Bool := false;   // Manual mode
      S_SEL : Int := 0;   // Select step to be output to S_NO
      S_ON : Bool := false;   // Activate step indicated in S_NO
      S_OFF : Bool := false;   // Deactivate step indicated S_NO
      T_PUSH : Bool := false;   // Enable transition to switch in semi automatic mode
   END_VAR
   VAR_OUTPUT
      S_NO : Int := 0;   // Step number
      S_MORE : Bool := false;   // More steps are available and can be shown in S_NO
      S_ACTIVE : Bool := false;   // Step indicated in S_NO is active
      ERR_FLT : Bool := false;   // Interlock or supervision group error
      AUTO_ON : Bool := false;   // Automatic mode is active
      TAP_ON : Bool := false;   // Semiautomatic mode/step with transition enabled
      TOP_ON : Bool := false;   // Semiautomatic mode/ignore transition enabled
      MAN_ON : Bool := false;   // Manual mode is active
   END_VAR
   VAR
      HMI_INFO : Array[0..8] of UInt;
      IF_PAR : G7_IfParPlus_V6;
      RT_DATA : G7_RTDataPlus_V6;   // Internal data area
      Trans1 : G7_TransitionPlus_V6;   // Transition structure
      Trans2 : G7_TransitionPlus_V6;   // Transition structure
      Trans3 : G7_TransitionPlus_V6;   // Transition structure
      Trans4 : G7_TransitionPlus_V6;   // Transition structure
      Trans5 : G7_TransitionPlus_V6;   // Transition structure
      Trans6 : G7_TransitionPlus_V6;   // Transition structure
      Trans7 : G7_TransitionPlus_V6;   // Transition structure
      Trans8 : G7_TransitionPlus_V6;   // Transition structure
      Trans9 : G7_TransitionPlus_V6;   // Transition structure
      Trans10 : G7_TransitionPlus_V6;   // Transition structure
      Trans11 : G7_TransitionPlus_V6;   // Transition structure
      Trans13 : G7_TransitionPlus_V6;   // Transition structure
      Trans14 : G7_TransitionPlus_V6;   // Transition structure
      Trans16 : G7_TransitionPlus_V6;   // Transition structure
      Trans17 : G7_TransitionPlus_V6;   // Transition structure
      Trans19 : G7_TransitionPlus_V6;   // Transition structure
      Trans20 : G7_TransitionPlus_V6;   // Transition structure
      Trans21 : G7_TransitionPlus_V6;   // Transition structure
      Step1 : G7_StepPlus_V6;   // Step structure
      Step2 : G7_StepPlus_V6;   // Step structure
      Step3 : G7_StepPlus_V6;   // Step structure
      Step4 : G7_StepPlus_V6;   // Step structure
      Step5 : G7_StepPlus_V6;   // Step structure
      Step6 : G7_StepPlus_V6;   // Step structure
      Step8 : G7_StepPlus_V6;   // Step structure
      Step9 : G7_StepPlus_V6;   // Step structure
      Step10 : G7_StepPlus_V6;   // Step structure
      Step12 : G7_StepPlus_V6;   // Step structure
      Step13 : G7_StepPlus_V6;   // Step structure
      Step14 : G7_StepPlus_V6;   // Step structure
      Step15 : G7_StepPlus_V6;   // Step structure
      Step16 : G7_StepPlus_V6;   // Step structure
      SINI : Array[0..1] of USInt;
      LSTT : Array[0..17] of USInt;
      ATAJ : Array[0..17] of USInt;
      ATAB : Array[0..17] of USInt;
      PSTT : Array[0..17] of USInt;
      NSTT : Array[0..17] of USInt;
      ASSJ : Array[0..13] of USInt;
      ASSB : Array[0..13] of USInt;
      PTTS : Array[0..13] of USInt;
      NTTS : Array[0..13] of USInt;
      SW_SQTS : Array[0..13] of USInt;
      SWITCH : Array[0..10] of USInt;
      TVX : Array[0..8] of USInt;
      TTX : Array[0..8] of USInt;
      TSX : Array[0..1] of USInt;
      S00X : Array[0..1] of USInt;
      SOFFX : Array[0..1] of USInt;
      SONX : Array[0..1] of USInt;
      SAX : Array[0..1] of USInt;
      SERRX : Array[0..14] of USInt;
      SMX : Array[0..14] of USInt;
      S0X : Array[0..14] of USInt;
      S1X : Array[0..14] of USInt;
      IL_ALARM_INST : Diag_Alarm;
      SUP_ALARM_INST : Diag_Alarm;
      STEP_TIME_ALARM_INST : Diag_Alarm;
      IEC_TIMER_INST : IEC_TIMER;
      TRANSACTION_FLAG : Bool := false;
   END_VAR
   // LSTT[13] := 255;
   // SINI[0] := 2;
   // LSTT[0] := 255;
   // LSTT[1] := 255;
   // LSTT[2] := 255;
   // LSTT[3] := 255;
   // LSTT[4] := 255;
   // LSTT[5] := 255;
   // LSTT[6] := 255;
   // LSTT[7] := 255;
   // LSTT[8] := 255;
   // LSTT[9] := 255;
   // LSTT[10] := 255;
   // ATAJ[1] := 1;
   // ATAJ[2] := 2;
   // ATAJ[3] := 3;
   // ATAJ[4] := 4;
   // ATAJ[5] := 6;
   // ATAJ[6] := 10;
   // ATAJ[7] := 7;
   // ATAJ[8] := 8;
   // ATAJ[9] := 9;
   // ATAJ[10] := 5;
   // ATAJ[11] := 11;
   // ATAJ[12] := 12;
   // ATAB[0] := 1;
   // ATAB[1] := 2;
   // ATAB[3] := 12;
   // ATAB[4] := 15;
   // ATAB[5] := 5;
   // ATAB[6] := 6;
   // ATAB[7] := 7;
   // ATAB[8] := 8;
   // ATAB[9] := 9;
   // ATAB[10] := 10;
   // ATAB[11] := 11;
   // ATAB[12] := 3;
   // PSTT[0] := 8;
   // PSTT[1] := 8;
   // PSTT[2] := 8;
   // PSTT[3] := 1;
   // PSTT[4] := 2;
   // PSTT[5] := 3;
   // PSTT[6] := 4;
   // PSTT[8] := 6;
   // PSTT[9] := 7;
   // PSTT[10] := 5;
   // PSTT[11] := 10;
   // PSTT[12] := 1;
   // NSTT[13] := 11;
   // NSTT[0] := 1;
   // NSTT[1] := 2;
   // NSTT[2] := 3;
   // NSTT[3] := 4;
   // NSTT[4] := 5;
   // NSTT[5] := 10;
   // NSTT[6] := 10;
   // NSTT[7] := 6;
   // NSTT[8] := 7;
   // NSTT[9] := 8;
   // NSTT[10] := 10;
   // ASSJ[1] := 1;
   // ASSJ[2] := 2;
   // ASSJ[3] := 3;
   // ASSJ[4] := 4;
   // ASSJ[5] := 5;
   // ASSJ[6] := 6;
   // ASSJ[7] := 7;
   // ASSJ[8] := 8;
   // ASSJ[9] := 9;
   // ASSJ[10] := 10;
   // ASSB[1] := 1;
   // ASSB[2] := 2;
   // ASSB[3] := 3;
   // ASSB[4] := 4;
   // ASSB[5] := 5;
   // ASSB[6] := 6;
   // ASSB[7] := 7;
   // ASSB[8] := 8;
   // ASSB[9] := 9;
   // ASSB[10] := 10;
   // PTTS[0] := 255;
   // PTTS[2] := 1;
   // PTTS[3] := 2;
   // PTTS[4] := 3;
   // PTTS[5] := 4;
   // PTTS[6] := 7;
   // PTTS[7] := 8;
   // PTTS[8] := 9;
   // PTTS[9] := 12;
   // PTTS[10] := 6;
   // NTTS[0] := 7;
   // NTTS[1] := 3;
   // NTTS[2] := 4;
   // NTTS[3] := 5;
   // NTTS[4] := 6;
   // NTTS[5] := 10;
   // NTTS[6] := 8;
   // NTTS[7] := 9;
   // NTTS[9] := 13;
   // NTTS[10] := 11;
   // SW_SQTS[1] := 1;
   // SW_SQTS[2] := 2;
   // SW_SQTS[3] := 3;
   // SW_SQTS[4] := 4;
   // SW_SQTS[5] := 5;
   // SW_SQTS[9] := 6;
   // SW_SQTS[10] := 7;
   // TVX[0] := 16#1;
   // TTX[0] := 16#1;
   // TSX[0] := 16#1;
   // S00X[0] := 16#1;
   // SOFFX[0] := 16#1;
   // SONX[0] := 16#1;
   // SAX[0] := 16#1;
   // SERRX[0] := 16#1;
   // SMX[0] := 16#1;
   // S0X[0] := 16#1;
   // S1X[0] := 16#1;
   // LSTT[12] := 255;
   // LSTT[14] := 4;
   // LSTT[15] := 255;
   // ATAJ[13] := 13;
   // ATAJ[14] := 14;
   // ATAJ[15] := 15;
   // ATAB[13] := 13;
   // ATAB[14] := 14;
   // ATAB[15] := 4;
   // PSTT[13] := 9;
   // PSTT[14] := 11;
   // PSTT[15] := 2;
   // NSTT[12] := 9;
   // NSTT[14] := 4;
   // NSTT[15] := 12;
   // ASSJ[11] := 11;
   // ASSJ[12] := 12;
   // ASSB[11] := 11;
   // ASSB[12] := 12;
   // PTTS[11] := 13;
   // PTTS[12] := 15;
   // NTTS[11] := 14;
   // NTTS[12] := 16;
   // SW_SQTS[11] := 6;
   // SW_SQTS[12] := 8;
   // LSTT[16] := 255;
   // LSTT[17] := 4;
   // ATAJ[16] := 16;
   // ATAJ[17] := 17;
   // ATAB[16] := 16;
   // ATAB[17] := 17;
   // PSTT[16] := 12;
   // PSTT[17] := 13;
   // NSTT[16] := 13;
   // NSTT[17] := 4;
   // ASSJ[13] := 13;
   // ASSB[13] := 13;
   // PTTS[13] := 16;
   // NTTS[13] := 17;
   // SW_SQTS[13] := 8;
BEGIN
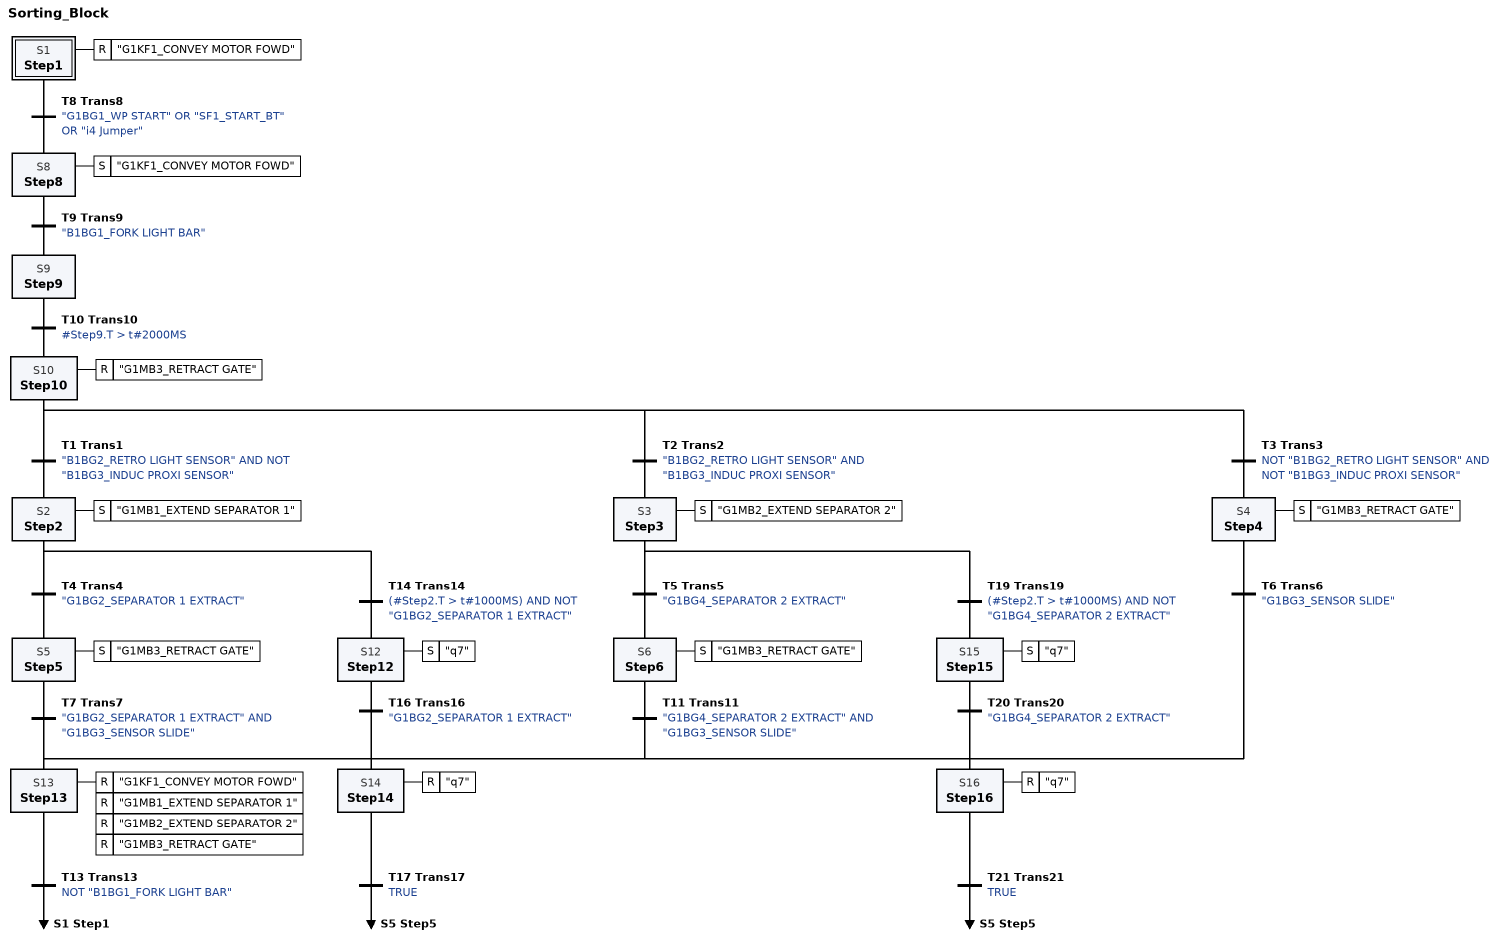
   // sequencer 1
   INITIAL_STEP Step1:   // S1, max time T#10S, warning time T#7S
              R    "G1KF1_CONVEY MOTOR FOWD"
   END_STEP
   TRANSITION Trans8 FROM Step1 TO Step8   // T8
      := "G1BG1_WP START" OR "SF1_START_BT" OR "i4 Jumper";
   END_TRANSITION
   STEP Step2:   // S2, max time T#10S, warning time T#7S
              S    "G1MB1_EXTEND SEPARATOR 1"
   END_STEP
   TRANSITION Trans4 FROM Step2 TO Step5   // T4
      := "G1BG2_SEPARATOR 1 EXTRACT";
   END_TRANSITION
   TRANSITION Trans14 FROM Step2 TO Step12   // T14
      := (#Step2.T > t#1000MS) AND NOT "G1BG2_SEPARATOR 1 EXTRACT";
   END_TRANSITION
   STEP Step3:   // S3, max time T#10S, warning time T#7S
              S    "G1MB2_EXTEND SEPARATOR 2"
   END_STEP
   TRANSITION Trans5 FROM Step3 TO Step6   // T5
      := "G1BG4_SEPARATOR 2 EXTRACT";
   END_TRANSITION
   TRANSITION Trans19 FROM Step3 TO Step15   // T19
      := (#Step2.T > t#1000MS) AND NOT "G1BG4_SEPARATOR 2 EXTRACT";
   END_TRANSITION
   STEP Step4:   // S4, max time T#10S, warning time T#7S
              S    "G1MB3_RETRACT GATE"
   END_STEP
   TRANSITION Trans6 FROM Step4 TO Step13   // T6
      := "G1BG3_SENSOR SLIDE";
   END_TRANSITION
   STEP Step5:   // S5, max time T#10S, warning time T#7S
              S    "G1MB3_RETRACT GATE"
   END_STEP
   TRANSITION Trans7 FROM Step5 TO Step13   // T7
      := "G1BG2_SEPARATOR 1 EXTRACT" AND "G1BG3_SENSOR SLIDE";
   END_TRANSITION
   STEP Step6:   // S6, max time T#10S, warning time T#7S
              S    "G1MB3_RETRACT GATE"
   END_STEP
   TRANSITION Trans11 FROM Step6 TO Step13   // T11
      := "G1BG4_SEPARATOR 2 EXTRACT" AND "G1BG3_SENSOR SLIDE";
   END_TRANSITION
   STEP Step8:   // S8, max time T#10S, warning time T#7S
              S    "G1KF1_CONVEY MOTOR FOWD"
   END_STEP
   TRANSITION Trans9 FROM Step8 TO Step9   // T9
      := "B1BG1_FORK LIGHT BAR";
   END_TRANSITION
   STEP Step10:   // S10, max time T#10S, warning time T#7S
              R    "G1MB3_RETRACT GATE"
   END_STEP
   TRANSITION Trans1 FROM Step10 TO Step2   // T1
      := "B1BG2_RETRO LIGHT SENSOR" AND NOT "B1BG3_INDUC PROXI SENSOR";
   END_TRANSITION
   TRANSITION Trans2 FROM Step10 TO Step3   // T2
      := "B1BG2_RETRO LIGHT SENSOR" AND "B1BG3_INDUC PROXI SENSOR";
   END_TRANSITION
   TRANSITION Trans3 FROM Step10 TO Step4   // T3
      := NOT "B1BG2_RETRO LIGHT SENSOR" AND NOT "B1BG3_INDUC PROXI SENSOR";
   END_TRANSITION
   STEP Step9:   // S9, max time T#10S, warning time T#7S
   END_STEP
   TRANSITION Trans10 FROM Step9 TO Step10   // T10
      := #Step9.T > t#2000MS;
   END_TRANSITION
   STEP Step12:   // S12, max time T#10S, warning time T#7S
              S    "q7"
   END_STEP
   TRANSITION Trans16 FROM Step12 TO Step14   // T16
      := "G1BG2_SEPARATOR 1 EXTRACT";
   END_TRANSITION
   STEP Step14:   // S14, max time T#10S, warning time T#7S
              R    "q7"
   END_STEP
   TRANSITION Trans17 FROM Step14 TO Step5   // T17, jump
      := TRUE;
   END_TRANSITION
   STEP Step15:   // S15, max time T#10S, warning time T#7S
              S    "q7"
   END_STEP
   TRANSITION Trans20 FROM Step15 TO Step16   // T20
      := "G1BG4_SEPARATOR 2 EXTRACT";
   END_TRANSITION
   STEP Step16:   // S16, max time T#10S, warning time T#7S
              R    "q7"
   END_STEP
   TRANSITION Trans21 FROM Step16 TO Step5   // T21, jump
      := TRUE;
   END_TRANSITION
   STEP Step13:   // S13, max time T#10S, warning time T#7S
              R    "G1KF1_CONVEY MOTOR FOWD"
              R    "G1MB1_EXTEND SEPARATOR 1"
              R    "G1MB2_EXTEND SEPARATOR 2"
              R    "G1MB3_RETRACT GATE"
   END_STEP
   TRANSITION Trans13 FROM Step13 TO Step1   // T13, jump
      := NOT "B1BG1_FORK LIGHT BAR";
   END_TRANSITION
END_FUNCTION_BLOCK

ORGANIZATION_BLOCK "Sorting_Main"   // OB1, LAD, ProgramCycle
TITLE = "Main Program Sweep (Cycle)"
{ S7_Optimized_Access := 'TRUE' }
VERSION : 0.1
   VAR_INPUT
      Initial_Call : Bool;   // Initial call of this OB
      Remanence : Bool;   // =True, if remanent data are available
   END_VAR
BEGIN

REGION Network 1
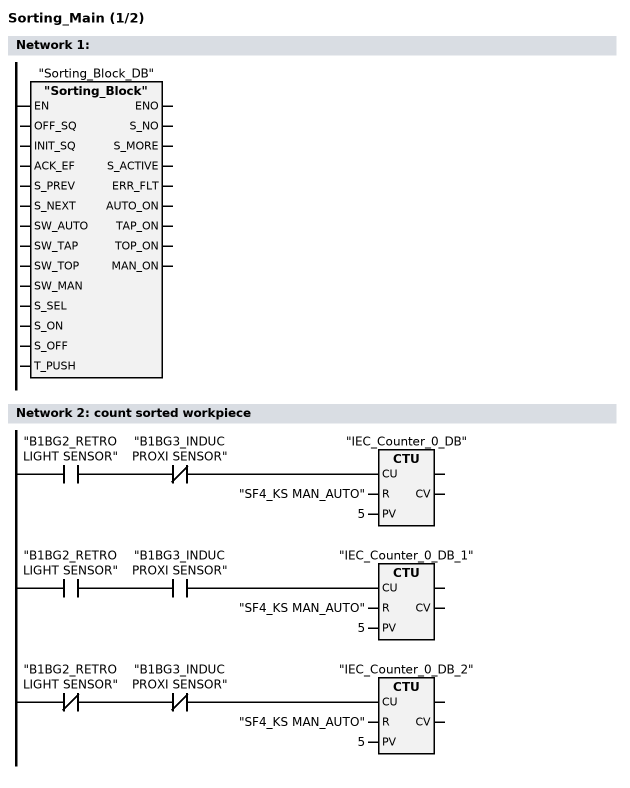
   RUNG wire#powerrail
      "Sorting_Block_DB"(OFF_SQ :=, INIT_SQ :=, ACK_EF :=, S_PREV :=, S_NEXT :=, SW_AUTO :=, SW_TAP :=, SW_TOP :=, SW_MAN :=, S_SEL :=, S_ON :=, S_OFF :=, T_PUSH :=, S_NO =>, S_MORE =>, S_ACTIVE =>, ERR_FLT =>, AUTO_ON =>, TAP_ON =>, TOP_ON =>, MAN_ON =>)
   END_RUNG
   // the same network as SCL:
   "Sorting_Block_DB"();   // "Sorting_Block"
END_REGION

REGION Network 2: count sorted workpiece
   "IEC_Counter_0_DB".CTU(CU := "B1BG2_RETRO LIGHT SENSOR" AND NOT "B1BG3_INDUC PROXI SENSOR",
                          R := "SF4_KS MAN_AUTO",
                          PV := 5);
   "IEC_Counter_0_DB_1".CTU(CU := "B1BG2_RETRO LIGHT SENSOR" AND "B1BG3_INDUC PROXI SENSOR",
                           R := "SF4_KS MAN_AUTO",
                           PV := 5);
   "IEC_Counter_0_DB_2".CTU(CU := NOT "B1BG2_RETRO LIGHT SENSOR" AND NOT "B1BG3_INDUC PROXI SENSOR",
                           R := "SF4_KS MAN_AUTO",
                           PV := 5);
END_REGION

REGION Network 3: reset
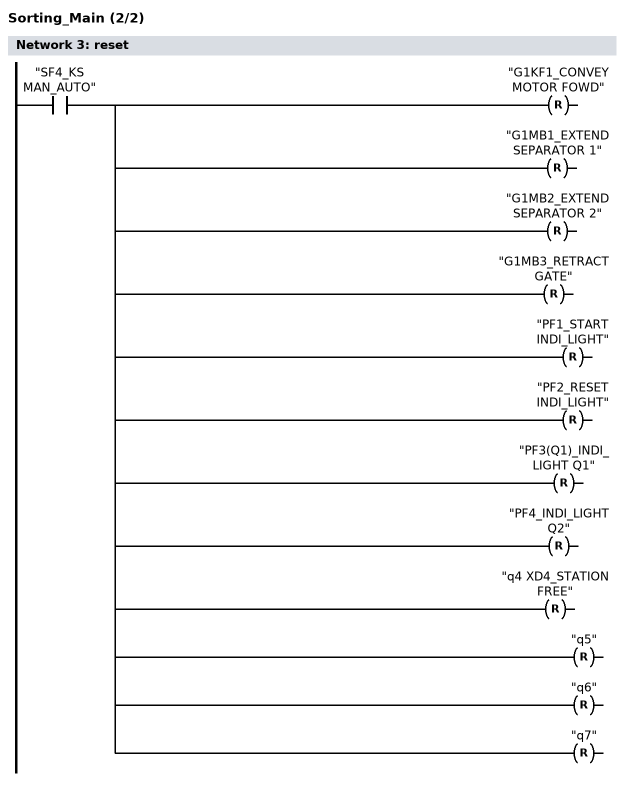
   RUNG wire#powerrail
      Contact( "SF4_KS MAN_AUTO" )
      wire#w1
      R_Coil( "G1KF1_CONVEY MOTOR FOWD" )
   END_RUNG
   RUNG wire#w1
      R_Coil( "G1MB1_EXTEND SEPARATOR 1" )
   END_RUNG
   RUNG wire#w1
      R_Coil( "G1MB2_EXTEND SEPARATOR 2" )
   END_RUNG
   RUNG wire#w1
      R_Coil( "G1MB3_RETRACT GATE" )
   END_RUNG
   RUNG wire#w1
      R_Coil( "PF1_START INDI_LIGHT" )
   END_RUNG
   RUNG wire#w1
      R_Coil( "PF2_RESET INDI_LIGHT" )
   END_RUNG
   RUNG wire#w1
      R_Coil( "PF3(Q1)_INDI_LIGHT Q1" )
   END_RUNG
   RUNG wire#w1
      R_Coil( "PF4_INDI_LIGHT Q2" )
   END_RUNG
   RUNG wire#w1
      R_Coil( "q4 XD4_STATION FREE" )
   END_RUNG
   RUNG wire#w1
      R_Coil( "q5" )
   END_RUNG
   RUNG wire#w1
      R_Coil( "q6" )
   END_RUNG
   RUNG wire#w1
      R_Coil( "q7" )
   END_RUNG
   // the same network as SCL:
   IF "SF4_KS MAN_AUTO" THEN
       "G1KF1_CONVEY MOTOR FOWD" := FALSE;
       "G1MB1_EXTEND SEPARATOR 1" := FALSE;
       "G1MB2_EXTEND SEPARATOR 2" := FALSE;
       "G1MB3_RETRACT GATE" := FALSE;
       "PF1_START INDI_LIGHT" := FALSE;
       "PF2_RESET INDI_LIGHT" := FALSE;
       "PF3(Q1)_INDI_LIGHT Q1" := FALSE;
       "PF4_INDI_LIGHT Q2" := FALSE;
       "q4 XD4_STATION FREE" := FALSE;
       "q5" := FALSE;
       "q6" := FALSE;
       "q7" := FALSE;
   END_IF;
END_REGION
END_ORGANIZATION_BLOCK